Universal Robots PolyScope program: nhom2_main.urp

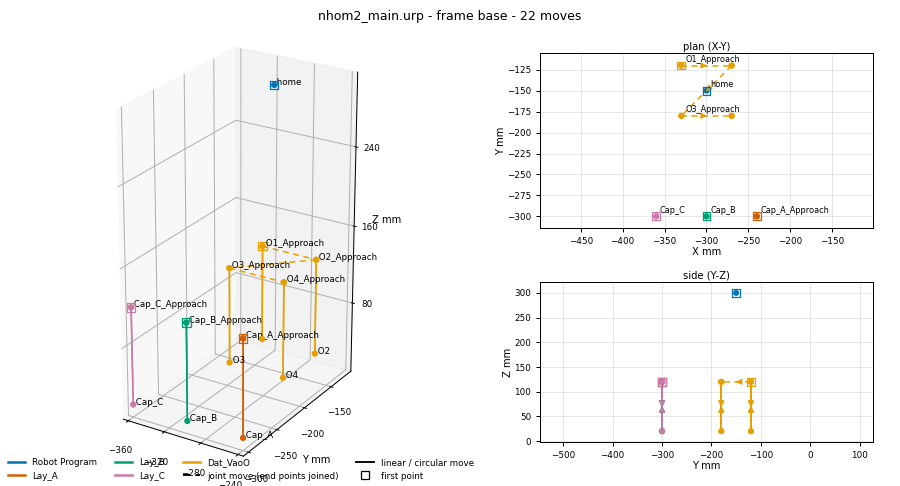
[picture p0: tool path of nhom2_main.urp in frame base, 22 of 22 moves have a stored position in this frame; points joined in program order, loops and branches not executed]
Program nhom2_main (installation=nhom2 directory=/home/ur/ursim-current/programs/Nhom2_CuoiKy createdIn=3.15.6.106324 lastSavedIn=3.15.6.106324 robotSerialNumber=2018339999)
Calibrated DH parameters: a=[0, -0.24365, -0.21325, 0, 0, 0]; d=[0.1519, 0, 0, 0.11235, 0.08535, 0.0819]; alpha=[1.570796, 0, 0, 1.570796, -1.570796, 0]; deltaTheta=[0, 0, 0, 0, 0, 0]
Robot Program (runOnlyOnce=true)
  ip := "192.168.61.1"
  n_read := 0
  rid := 0
  ok := False
  okk := False
  st := 0
  cls := 0
  slot := 0
  conf := 0.0
  n_dat := 0
  n_khay_xong := 0
  n_cho := 0
  n_loi := 0
  retries := 0
  msg := ""
  chay := True
  Set DigitalOutput pin=digital_out[0]; digitalValue=0
  Set DigitalOutput pin=digital_out[1]; digitalValue=0
  Set DigitalOutput pin=digital_out[2]; digitalValue=0
  MoveJ speed 60 deg/s, acceleration 80 deg/s^2 (useActiveTCP=true)
    Waypoint home: TCP in base x=-300 y=-150 z=300 mm, rx=-3.1412 ry=0 rz=0 rad; joints [7.008, -81.262, 56.541, -65.276, -90.023, 97.008] deg; flange x=-300 y=-150.041 z=400 mm, rx=-3.1412 ry=0 rz=0 rad
  Script: okk = socket_open(ip, 5000, "py")
  Popup Message (haltProgram=false message=okk inputType=Variable) variable=okk
  cid := 0
  r := [0,0,0,0,0,0,0,0,0]
  Loop While (checkContinuously=false) expression=chay == True
    cid := cid + 1
    ok := False
    Script: socket_send_line(str_cat("GET,", to_str(cid)), "py")
    Script: r = socket_read_ascii_float(8, "py", 5)
    Script: n_read = r[0]
    If n_read == 8
      Script: rid = r[1]
      If rid == cid
        Script: st = r[2]
        Script: cls = r[3]
        Script: conf = r[7]
        Script: slot = r[8]
        ok := True
    If ok == False
      Set DigitalOutput pin=digital_out[1]; digitalValue=1
      n_loi := n_loi + 1
      Script: socket_close("py")
      Wait Sleep waitTime=1
      Script: okk = socket_open(ip, 5000, "py")
      retries := retries + 1
      If retries >= 5
        Popup Message (haltProgram=false message=Mat ket noi, kiem tra bridge inputType=Text)
        chay := False
    ElseIf st == 1 and conf >= 0.5 and ((cls==1 and (slot==1 or slot==2)) or (cls==2 and slot==3) or (cls==3 and slot==4))
      Set DigitalOutput pin=digital_out[1]; digitalValue=0
      retries := 0
      If cls == 1
        Call Lay_A
      ElseIf cls == 2
        Call Lay_B
      ElseIf cls == 3
        Call Lay_C
      Call Dat_VaoO
      Script: socket_send_line(str_cat("DONE,", to_str(cid)), "py")
      n_dat := n_dat + 1
      Set DigitalOutput pin=digital_out[2]; digitalValue=1
      Wait Sleep waitTime=0.2
      Set DigitalOutput pin=digital_out[2]; digitalValue=0
    ElseIf st == 3
      Set DigitalOutput pin=digital_out[1]; digitalValue=0
      Script: socket_send_line(str_cat("DONE,", to_str(cid)), "py")
      n_khay_xong := n_khay_xong + 1
      chay := False
    Else 
      n_cho := n_cho + 1
      retries := retries + 1
      Wait Sleep waitTime=0.5
      If retries >= 3
        Popup Message (haltProgram=true message=Can nguoi van hanh kiem tra inputType=Text)
        chay := False
  Script: msg = str_cat("n_dat=", str_cat(to_str(n_dat), str_cat("  n_khay_xong=", str_cat(to_str(n_khay_xong), str_cat("  n_cho=", str_cat(to_str(n_cho), str_cat("  n_loi=", to_str(n_loi))))))))
  Popup Message (haltProgram=false inputType=Variable) variable=msg
  Script: socket_close("py")
SubProgram -> Lay_A
SubProgram -> Lay_B
SubProgram -> Lay_C
SubProgram -> Dat_VaoO
SubProgram Lay_A (keepSynchronizedWithDisk=false)
  MoveJ speed 60 deg/s, acceleration 80 deg/s^2 (useActiveTCP=true)
    Waypoint Cap_A_Approach: TCP in base x=-240 y=-300 z=120 mm, rx=-3.1412 ry=0 rz=0 rad; joints [34.346, -69.854, 91.518, -111.651, -90.019, 124.346] deg; flange x=-240 y=-300.041 z=220 mm, rx=-3.1412 ry=0 rz=0 rad
  MoveL speed 250 mm/s, acceleration 1200 mm/s^2 (useActiveTCP=true) feature=Base
    Waypoint Cap_A: TCP in base x=-240 y=-300 z=20 mm, rx=-3.1412 ry=0 rz=0 rad; joints [-111.652, -123.37, -102.649, -44.003, 89.991, -201.652] deg; flange x=-240 y=-300.041 z=120 mm, rx=-3.1412 ry=0 rz=0 rad
  Set DigitalOutput pin=digital_out[0]; digitalValue=1
  Wait Sleep waitTime=0.5
  MoveL speed 250 mm/s, acceleration 1200 mm/s^2 (useActiveTCP=true) feature=Base
    Waypoint Cap_A_Approach: TCP in base x=-240 y=-300 z=120 mm, rx=-3.1412 ry=0 rz=0 rad; joints [34.346, -69.854, 91.518, -111.651, -90.019, 124.346] deg; flange x=-240 y=-300.041 z=220 mm, rx=-3.1412 ry=0 rz=0 rad
SubProgram Lay_B (keepSynchronizedWithDisk=false)
  MoveJ speed 60 deg/s, acceleration 80 deg/s^2 (useActiveTCP=true)
    Waypoint Cap_B_Approach: TCP in base x=-300 y=-300 z=120 mm, rx=-3.1412 ry=0 rz=0 rad; joints [29.653, -60.542, 77.481, -106.928, -90.02, 119.653] deg; flange x=-300 y=-300.041 z=220 mm, rx=-3.1412 ry=0 rz=0 rad
  MoveL speed 250 mm/s, acceleration 1200 mm/s^2 (useActiveTCP=true) feature=Base
    Waypoint Cap_B: TCP in base x=-300 y=-300 z=20 mm, rx=-3.1412 ry=0 rz=0 rad; joints [-119.639, -130.628, -88.609, -50.783, 89.988, -209.639] deg; flange x=-300 y=-300.041 z=120 mm, rx=-3.1412 ry=0 rz=0 rad
  Set DigitalOutput pin=digital_out[0]; digitalValue=1
  Wait Sleep waitTime=0.5
  MoveL speed 250 mm/s, acceleration 1200 mm/s^2 (useActiveTCP=true) feature=Base
    Waypoint Cap_B_Approach: TCP in base x=-300 y=-300 z=120 mm, rx=-3.1412 ry=0 rz=0 rad; joints [29.653, -60.542, 77.481, -106.928, -90.02, 119.653] deg; flange x=-300 y=-300.041 z=220 mm, rx=-3.1412 ry=0 rz=0 rad
SubProgram Lay_C (keepSynchronizedWithDisk=false)
  MoveJ speed 60 deg/s, acceleration 80 deg/s^2 (useActiveTCP=true)
    Waypoint Cap_C_Approach: TCP in base x=-360 y=-300 z=120 mm, rx=-3.1412 ry=0 rz=0 rad; joints [25.942, -49.203, 58.496, -99.283, -90.021, 115.942] deg; flange x=-360 y=-300.041 z=220 mm, rx=-3.1412 ry=0 rz=0 rad
  MoveL speed 250 mm/s, acceleration 1200 mm/s^2 (useActiveTCP=true) feature=Base
    Waypoint Cap_C: TCP in base x=-360 y=-300 z=20 mm, rx=-3.1412 ry=0 rz=0 rad; joints [-126.317, -139.633, -70.727, -59.66, 89.986, -216.317] deg; flange x=-360 y=-300.041 z=120 mm, rx=-3.1412 ry=0 rz=0 rad
  Set DigitalOutput pin=digital_out[0]; digitalValue=1
  Wait Sleep waitTime=0.5
  MoveL speed 250 mm/s, acceleration 1200 mm/s^2 (useActiveTCP=true) feature=Base
    Waypoint Cap_C_Approach: TCP in base x=-360 y=-300 z=120 mm, rx=-3.1412 ry=0 rz=0 rad; joints [25.942, -49.203, 58.496, -99.283, -90.021, 115.942] deg; flange x=-360 y=-300.041 z=220 mm, rx=-3.1412 ry=0 rz=0 rad
SubProgram Dat_VaoO (keepSynchronizedWithDisk=false)
  If slot == 1
    MoveJ speed 60 deg/s, acceleration 80 deg/s^2 (useActiveTCP=true)
      Waypoint O1_Approach: TCP in base x=-330 y=-120 z=120 mm, rx=-3.1412 ry=0 rz=0 rad; joints [1.336, -77.43, 101.746, -114.315, -90.023, 91.336] deg; flange x=-330 y=-120.041 z=220 mm, rx=-3.1412 ry=0 rz=0 rad
    MoveL speed 250 mm/s, acceleration 1200 mm/s^2 (useActiveTCP=true) feature=Base
      Waypoint O1: TCP in base x=-330 y=-120 z=20 mm, rx=-3.1412 ry=0 rz=0 rad; joints [-141.347, -117.679, -113.329, -39.006, 89.982, -231.347] deg; flange x=-330 y=-120.041 z=120 mm, rx=-3.1412 ry=0 rz=0 rad
    Set DigitalOutput pin=digital_out[0]; digitalValue=0
    Wait Sleep waitTime=0.5
    MoveL speed 250 mm/s, acceleration 1200 mm/s^2 (useActiveTCP=true) feature=Base
      Waypoint O1_Approach: TCP in base x=-330 y=-120 z=120 mm, rx=-3.1412 ry=0 rz=0 rad; joints [1.336, -77.43, 101.746, -114.315, -90.023, 91.336] deg; flange x=-330 y=-120.041 z=220 mm, rx=-3.1412 ry=0 rz=0 rad
  ElseIf slot == 2
    MoveJ speed 60 deg/s, acceleration 80 deg/s^2 (useActiveTCP=true)
      Waypoint O2_Approach: TCP in base x=-270 y=-120 z=120 mm, rx=-3.1412 ry=0 rz=0 rad; joints [1.629, -90.857, 116.899, -116.041, -90.023, 91.629] deg; flange x=-270 y=-120.041 z=220 mm, rx=-3.1412 ry=0 rz=0 rad
    MoveL speed 250 mm/s, acceleration 1200 mm/s^2 (useActiveTCP=true) feature=Base
      Waypoint O2: TCP in base x=-270 y=-120 z=20 mm, rx=-3.1412 ry=0 rz=0 rad; joints [-133.678, -108.167, -130.155, -31.695, 89.984, -223.678] deg; flange x=-270 y=-120.041 z=120 mm, rx=-3.1412 ry=0 rz=0 rad
    Set DigitalOutput pin=digital_out[0]; digitalValue=0
    Wait Sleep waitTime=0.5
    MoveL speed 250 mm/s, acceleration 1200 mm/s^2 (useActiveTCP=true) feature=Base
      Waypoint O2_Approach: TCP in base x=-270 y=-120 z=120 mm, rx=-3.1412 ry=0 rz=0 rad; joints [1.629, -90.857, 116.899, -116.041, -90.023, 91.629] deg; flange x=-270 y=-120.041 z=220 mm, rx=-3.1412 ry=0 rz=0 rad
  ElseIf slot == 3
    MoveJ speed 60 deg/s, acceleration 80 deg/s^2 (useActiveTCP=true)
      Waypoint O3_Approach: TCP in base x=-330 y=-180 z=120 mm, rx=-3.1412 ry=0 rz=0 rad; joints [11.232, -71.752, 94.188, -112.432, -90.023, 101.232] deg; flange x=-330 y=-180.041 z=220 mm, rx=-3.1412 ry=0 rz=0 rad
    MoveL speed 250 mm/s, acceleration 1200 mm/s^2 (useActiveTCP=true) feature=Base
      Waypoint O3: TCP in base x=-330 y=-180 z=20 mm, rx=-3.1412 ry=0 rz=0 rad; joints [-133.991, -121.924, -105.396, -42.696, 89.984, -223.991] deg; flange x=-330 y=-180.041 z=120 mm, rx=-3.1412 ry=0 rz=0 rad
    Set DigitalOutput pin=digital_out[0]; digitalValue=0
    Wait Sleep waitTime=0.5
    MoveL speed 250 mm/s, acceleration 1200 mm/s^2 (useActiveTCP=true) feature=Base
      Waypoint O3_Approach: TCP in base x=-330 y=-180 z=120 mm, rx=-3.1412 ry=0 rz=0 rad; joints [11.232, -71.752, 94.188, -112.432, -90.023, 101.232] deg; flange x=-330 y=-180.041 z=220 mm, rx=-3.1412 ry=0 rz=0 rad
  ElseIf slot == 4
    MoveJ speed 60 deg/s, acceleration 80 deg/s^2 (useActiveTCP=true)
      Waypoint O4_Approach: TCP in base x=-270 y=-180 z=120 mm, rx=-3.1412 ry=0 rz=0 rad; joints [13.447, -83.681, 109.287, -115.6, -90.023, 103.447] deg; flange x=-270 y=-180.041 z=220 mm, rx=-3.1412 ry=0 rz=0 rad
    MoveL speed 250 mm/s, acceleration 1200 mm/s^2 (useActiveTCP=true) feature=Base
      Waypoint O4: TCP in base x=-270 y=-180 z=20 mm, rx=-3.1412 ry=0 rz=0 rad; joints [-126.045, -113.158, -121.517, -35.343, 89.986, -216.045] deg; flange x=-270 y=-180.041 z=120 mm, rx=-3.1412 ry=0 rz=0 rad
    Set DigitalOutput pin=digital_out[0]; digitalValue=0
    Wait Sleep waitTime=0.5
    MoveL speed 250 mm/s, acceleration 1200 mm/s^2 (useActiveTCP=true) feature=Base
      Waypoint O4_Approach: TCP in base x=-270 y=-180 z=120 mm, rx=-3.1412 ry=0 rz=0 rad; joints [13.447, -83.681, 109.287, -115.6, -90.023, 103.447] deg; flange x=-270 y=-180.041 z=220 mm, rx=-3.1412 ry=0 rz=0 rad
